Fanuc KAREL source: kb00022.KL

-- PROVISIONAL review KL for V770-1; original PC SHA256 2f76e62b3bb9fae372f9df83dc9d507489a7a13884a6f5a50a1521072ec68d21
-- Incomplete behavior may be omitted. Consult companion uncertainty JSON. Do not deploy.
PROGRAM KB00022
%NOLOCKGROUP
BEGIN
  -- UNRESOLVED_PC offsets 5-12; opcodes 9D,23
  -- UNRESOLVED_PC offsets 17-27; opcodes 27,22,31
  -- UNRESOLVED_PC offsets 32-36; opcodes 7F
END KB00022
